(*
SPDX-FileCopyrightText: © 2026 Oleksandr Tiutyk <trofimich@gmail.com>
SPDX-License-Identifier: MIT
License: https://opensource.org/license/mit
*)

(*!
<summary>Observes parent resource release without using a real resource.</summary>
<description>
Configure Child and ThrowOnStartRelease through SetChild and SetThrowOnStartRelease before the queue starts.
Child is borrowed and must outlive this manager. Acquisition takes one Execute; release takes two.
EarlyRelease records any request while Child is RUNNING. ReleaseCalls and EarlyRelease are observations only.
ResetFixture clears the synthetic state between independent test runs. No physical resource is created.
</description>
*)

FUNCTION_BLOCK QueueCleanupResource EXTENDS TOF_Core.Object IMPLEMENTS TOF_Core.IResourceManager
VAR_OUTPUT
	//! <summary>Borrowed child whose RUNNING state must prevent parent release.</summary>
	Child : TOF_Tasks.ITask;
	//! <summary>Raise a terminal release-attempt error on StartRelease.</summary>
	ThrowOnStartRelease : BOOL;
	//! <summary>Total StartRelease calls; read-only to tests.</summary>
	ReleaseCalls : UINT;
	//! <summary>Records whether release was requested while Child was RUNNING.</summary>
	EarlyRelease : BOOL;
END_VAR
VAR CONSTANT
	//! <summary>Execute calls required to complete synthetic release after its request.</summary>
	_ReleaseSteps : UINT := 2;
END_VAR
VAR_STAT
	//! <summary>Class name shared by all instances of this function block.</summary>
	_ClassName : STRING := __POUNAME();
END_VAR
VAR
	_Acquired : BOOL;
	_Acquiring : BOOL;
	_Releasing : BOOL;
	_ReleaseProgress : UINT;
END_VAR

{attribute 'monitoring' := 'call'}
PROPERTY ClassName : REFERENCE TO STRING
GET
ClassName REF= _ClassName;
END_GET
END_PROPERTY

(*!
<summary>Advances one synthetic acquisition or release step.</summary>
<description>
Idle calls do nothing; all operations are bounded and perform no I/O.
</description>
*)
METHOD Execute
IF _Acquiring THEN
	_Acquired := TRUE;
	_Acquiring := FALSE;
ELSIF _Releasing THEN
	_ReleaseProgress := _ReleaseProgress + 1;

	IF _ReleaseProgress >= _ReleaseSteps THEN
		_Acquired := FALSE;
		_Releasing := FALSE;
	END_IF
END_IF
END_METHOD

(*!
<summary>Returns this live fixture as the borrowed synthetic resource.</summary>
<description>
No real handle is created. The caller must not delete the returned object.
</description>
*)
METHOD GetResource : TOF_Core.IObject
GetResource := THIS^;
END_METHOD

(*!
<summary>Borrows the test library namespace.</summary>
*)

{attribute 'monitoring' := 'call'}
PROPERTY NamespaceName : REFERENCE TO STRING
GET
NamespaceName REF= CurrentNamespace.Name;
END_GET
END_PROPERTY

(*!
<summary>Reports whether the synthetic resource is held.</summary>
<description>
Has no side effects and does not throw.
</description>
*)

{attribute 'monitoring' := 'call'}
PROPERTY ResourceAcquired : BOOL
GET
ResourceAcquired := _Acquired;
END_GET
END_PROPERTY

(*!
<summary>Reports the concrete fixture size.</summary>
*)

{attribute 'monitoring' := 'call'}
PROPERTY SelfSize : ULINT
GET
SelfSize := XSIZEOF(THIS^);
END_GET
END_PROPERTY

(*!
<summary>Restores an idle synthetic resource and clears its observations.</summary>
<description>
Call only after the owning queue and children have stopped or before they start. Keeps the borrowed child
binding. Clears simulated state even after an injected terminal release error. Performs no physical release.
</description>
*)
METHOD INTERNAL ResetFixture
_Acquired := FALSE;
_Acquiring := FALSE;
_Releasing := FALSE;
_ReleaseProgress := 0;
ReleaseCalls := 0;
EarlyRelease := FALSE;
ThrowOnStartRelease := FALSE;
END_METHOD

(*!
<summary>Sets the child observed during resource release.</summary>
<description>
Call before the queue starts. The child is borrowed and must outlive the resource manager.
</description>
<param name="child">Child whose RUNNING state is observed during release.</param>
*)
METHOD INTERNAL SetChild
VAR_INPUT
	child : TOF_Tasks.ITask;
END_VAR
THIS^.Child := child;
END_METHOD

(*!
<summary>Configures the resource's release failure injection.</summary>
<description>
Call before the queue starts. Changes only the failure setting; resource progress and observations are
preserved.
</description>
<param name="throwOnStartRelease">Whether StartRelease raises the synthetic release-attempt error.</param>
*)
METHOD INTERNAL SetThrowOnStartRelease
VAR_INPUT
	throwOnStartRelease : BOOL;
END_VAR
THIS^.ThrowOnStartRelease := throwOnStartRelease;
END_METHOD

(*!
<summary>Requests synthetic acquisition completed by the next Execute.</summary>
<description>
Called once per acquire phase. Does nothing when already acquired.
</description>
*)
METHOD StartAcquire
IF NOT _Acquired THEN
	_Acquiring := TRUE;
END_IF
END_METHOD

(*!
<summary>Records release ordering and starts synthetic release.</summary>
<description>
Records EarlyRelease before optionally throwing. A thrown release deliberately leaves ResourceAcquired TRUE;
this models a failed terminal attempt without holding any real resource.
</description>
*)
METHOD StartRelease
VAR
	failure : TOF_Core.StandardException;
END_VAR
ReleaseCalls := ReleaseCalls + 1;

IF Child <> 0 AND_THEN Child.State.Running THEN
	EarlyRelease := TRUE;
END_IF

IF ThrowOnStartRelease THEN
	failure.Throw(
		sourceNamespaceName := NamespaceName,
		sourceClassName := ClassName,
		sourcePOUName := __POUNAME(),
		sourcePosition := __POSITION(),
		message := "Parent release failure"
	);
END_IF

_ReleaseProgress := 0;
_Releasing := TRUE;
END_METHOD

END_FUNCTION_BLOCK

(* stored: Version 1.1.0.1, ProductVersion 3.1.4026.21
   POU QueueCleanupResource: Id {a974a31d-e888-4192-a36d-7424fa95549f}, SpecialFunc None
   Folder Internal methods: Id {8c23ba67-ee83-413c-b94a-1f55ab5252ad}
   Property ClassName: Id {7786eeca-4512-4cfb-bcd5-b9e169863e53}
   Get Get: Id {d02f21ef-9ca8-4378-8d38-8cbd1eebf4bb}
   Method Execute: Id {1754ea46-b3bd-409b-85b9-07835c3639c1}
   Method GetResource: Id {43736e26-7196-40e1-9455-cadb39069ec9}
   Property NamespaceName: Id {3c9f5fc1-495b-4240-863e-f2c083b24cf8}
   Get Get: Id {4577d80a-1115-42ea-a888-c338c605846c}
   Property ResourceAcquired: Id {07ef79e6-8e33-4f3f-96bb-ccbaa770fbc6}
   Get Get: Id {ea6ac594-b94e-4c92-b4f5-1b226b4c9bcc}
   Property SelfSize: Id {0417d685-2ae3-4048-87c6-ee3c564ff270}
   Get Get: Id {876cfd53-2bbe-427e-a3c4-d370208b8741}
   Method ResetFixture: Id {6d8a0ca7-e1e0-4751-8923-72d4272f6f8d}
   Method SetChild: Id {860691b1-452d-4651-8e8f-fd8460ed6dd0}
   Method SetThrowOnStartRelease: Id {01b079c3-5180-4776-88bd-548796fd291e}
   Method StartAcquire: Id {b7a8d6be-c5a9-47a4-9209-6448343e8be2}
   Method StartRelease: Id {1529eda6-d75b-4f72-9327-20cbddf1bb98} *)
